{attribute 'qualified_only'}
{attribute 'strict'}
{attribute 'to_string'}
TYPE E_Request_List :
(
eNone :=0,
eDrain,

eCIP3,
eCIP5,



eWaterPrepare,
eDissolve,
eProduction,
eDisconnectTank,

eFinish
);
END_TYPE

(* stored: Version 1.1.0.1, ProductVersion 3.1.4024.12
   DUT E_Request_List: Id {c21fbe3a-d713-46bb-8806-9ab640ffc4cd} *)
